// TIA Portal V21 export
// export: Created 2026-10-14T03:11:19.8058014Z, ExportSetting WithDefaults, DisplayName Totally Integrated Automation Portal, DisplayVersion V21, DisplayName STEP 7 Professional, DisplayVersion V21, DisplayName STEP 7 Safety, DisplayVersion V21, DisplayName Tech WebApplication, DisplayVersion V21, DisplayName WinCC Basic/Comfort/Advanced, DisplayVersion V21, DisplayName WinCC Unified, DisplayVersion V21
TagTable "PID_Compact"
  PID_Compact_1_Input : Real  (HMI_Connection_1, 100 ms)
  PID_Compact_1_Output : Real  (HMI_Connection_1, 100 ms)
  PID_Compact_1_Setpoint : Real  (HMI_Connection_1, 100 ms)
  PID_Compact_1_Input_PER : Int  (HMI_Connection_1, 1 s)
  PID_Compact_1_Disturbance : Real  (HMI_Connection_1, 1 s)
  PID_Compact_1_ManualEnable : Bool  (HMI_Connection_1, 1 s)
  PID_Compact_1_ManualValue : Real  (HMI_Connection_1, 1 s)
  PID_Compact_1_ErrorAck : Bool  (HMI_Connection_1, 1 s)
  PID_Compact_1_Reset : Bool  (HMI_Connection_1, 1 s)
  PID_Compact_1_ModeActivate : Bool  (HMI_Connection_1, 1 s)
  PID_Compact_1_ScaledInput : Real  (HMI_Connection_1, 1 s)
  PID_Compact_1_Output_PER : Int  (HMI_Connection_1, 1 s)
  PID_Compact_1_Output_PWM : Bool  (HMI_Connection_1, 1 s)
  PID_Compact_1_SetpointLimit_H : Bool  (HMI_Connection_1, 1 s)
  PID_Compact_1_SetpointLimit_L : Bool  (HMI_Connection_1, 1 s)
  PID_Compact_1_InputWarning_H : Bool  (HMI_Connection_1, 1 s)
  PID_Compact_1_InputWarning_L : Bool  (HMI_Connection_1, 1 s)
  PID_Compact_1_State : Int  (HMI_Connection_1, 1 s)
  PID_Compact_1_Error : Bool  (HMI_Connection_1, 1 s)
  PID_Compact_1_ErrorBits : DWord  (HMI_Connection_1, 1 s)
  PID_Compact_1_Mode : Int  (HMI_Connection_1, 1 s)
  PID_Compact_1_InternalVersion : DWord  (HMI_Connection_1, 1 s)
  PID_Compact_1_IntegralResetMode : Int  (HMI_Connection_1, 1 s)
  PID_Compact_1_OverwriteInitialOutputValue : Real  (HMI_Connection_1, 1 s)
  PID_Compact_1_RunModeByStartup : Bool  (HMI_Connection_1, 1 s)
  PID_Compact_1_LoadBackUp : Bool  (HMI_Connection_1, 1 s)
  PID_Compact_1_SetSubstituteOutput : Bool  (HMI_Connection_1, 1 s)
  PID_Compact_1_PhysicalUnit : Int  (HMI_Connection_1, 1 s)
  PID_Compact_1_PhysicalQuantity : Int  (HMI_Connection_1, 1 s)
  PID_Compact_1_ActivateRecoverMode : Bool  (HMI_Connection_1, 1 s)
  PID_Compact_1_Warning : DWord  (HMI_Connection_1, 1 s)
  PID_Compact_1_WarningInternal : DWord  (HMI_Connection_1, 1 s)
  PID_Compact_1_Progress : Real  (HMI_Connection_1, 1 s)
  PID_Compact_1_CurrentSetpoint : Real  (HMI_Connection_1, 1 s)
  PID_Compact_1_CancelTuningLevel : Real  (HMI_Connection_1, 1 s)
  PID_Compact_1_SubstituteOutput : Real  (HMI_Connection_1, 1 s)
  PID_Compact_1_Config : PID_CompactConfig  (HMI_Connection_1, 1 s)
    TagStructureMember "InputPerOn"
    TagStructureMember "InvertControl"
    TagStructureMember "OutputSelect"
    TagStructureMember "InputUpperLimit"
    TagStructureMember "InputLowerLimit"
    TagStructureMember "InputUpperWarning"
    TagStructureMember "InputLowerWarning"
    TagStructureMember "OutputUpperLimit"
    TagStructureMember "OutputLowerLimit"
    TagStructureMember "SetpointUpperLimit"
    TagStructureMember "SetpointLowerLimit"
    TagStructureMember "MinimumOnTime"
    TagStructureMember "MinimumOffTime"
    TagStructureMember "InputScaling"
      TagStructureMember "UpperPointIn"
      TagStructureMember "LowerPointIn"
      TagStructureMember "UpperPointOut"
      TagStructureMember "LowerPointOut"
  PID_Compact_1_CycleTime : PID_CycleTime  (HMI_Connection_1, 1 s)
    TagStructureMember "StartEstimation"
    TagStructureMember "EnEstimation"
    TagStructureMember "EnMonitoring"
    TagStructureMember "Value"
  PID_Compact_1_CtrlParamsBackUp : PID_CompactControlParams  (HMI_Connection_1, 1 s)
    TagStructureMember "SetByUser"
    TagStructureMember "Gain"
    TagStructureMember "Ti"
    TagStructureMember "Td"
    TagStructureMember "TdFiltRatio"
    TagStructureMember "PWeighting"
    TagStructureMember "DWeighting"
    TagStructureMember "Cycle"
    TagStructureMember "DeadZone"
  PID_Compact_1_PIDSelfTune : PID_CompactSelfTune  (HMI_Connection_1, 1 s)
    TagStructureMember "SUT"
      TagStructureMember "CalculateParams"
      TagStructureMember "TuneRule"
      TagStructureMember "State"
    TagStructureMember "TIR"
      TagStructureMember "RunIn"
      TagStructureMember "CalculateParams"
      TagStructureMember "TuneRule"
      TagStructureMember "State"
  PID_Compact_1_PIDCtrl : PID_CompactControl  (HMI_Connection_1, 100 ms)
    TagStructureMember "PIDInit"
    TagStructureMember "IntegralSum"
  PID_Compact_1_Retain : PID_CompactRetain  (HMI_Connection_1, 1 s)
    TagStructureMember "CtrlParams"
      TagStructureMember "SetByUser"
      TagStructureMember "Gain"
      TagStructureMember "Ti"
      TagStructureMember "Td"
      TagStructureMember "TdFiltRatio"
      TagStructureMember "PWeighting"
      TagStructureMember "DWeighting"
      TagStructureMember "Cycle"
      TagStructureMember "DeadZone"
